(* IEC 61131-3 sources: Test-Git_ESME26/TestProgettoESME_26.fbsproj/TemplateFullProgrammingFramework_Migration.device.xml.v3^/Plc Logic.plclogic.xml.v3^/Application.application.xml.v3^/TemplateFullProgrammingFramework/Examples/ExampleDiagSources/FB_ApplicationLoggerDiagSource.fb.st^, 6 files *)

(* ---- CancelWriting.meth.st ---- *)
METHOD INTERNAL CancelWriting
VAR_INPUT
END_VAR

(* Deactivate writing if we are (for whatever reason) no longer adressed.
   May happen in case network connection with Diagnostics is disrupted or Source will be disabled *)

THIS^.diOldCmd			:= 0;
THIS^.diCmdExecState	:= 0;

(* ---- DiagQuit.meth.st ---- *)
METHOD INTERNAL DiagQuit
VAR_INPUT
END_VAR

IF THIS^.i_xEnable AND THIS^.q_xActive AND THIS^.q_etDiag <> GD.ET_Diag.Ok AND THIS^.diState = 0 THEN

	THIS^.rtrigDiagQuit(CLK := THIS^.i_xDiagQuit);
	IF THIS^.rtrigDiagQuit.Q THEN
		CancelWriting();

		THIS^.udiOwnSourceId	:= 0;

		THIS^.fbTreeWriter.FB_Init(bInitRetains := FALSE, bInCopyCode := FALSE);

		THIS^.q_xReady		:= TRUE;
		THIS^.q_etDiag		:= GD.ET_Diag.Ok;
		THIS^.q_etDiagExt	:= ET_DiagExt.WaitUntilDiagnosticsManagerReady;
		THIS^.q_sMsg		:= '';

		THIS^.diState := 10;
	END_IF

END_IF

(* ---- ExceptionDuringWriting.meth.st ---- *)
METHOD INTERNAL ExceptionDuringWriting : BOOL
VAR_INPUT
END_VAR

(* exception during writing *)
CASE THIS^.etDiagExtBufferTPL OF
	TPL.ET_DiagExt.TreeStartAlreadySuccessfullyCalled,		// FB_TreeWriter.TreeStart
	TPL.ET_DiagExt.FileIdNotSet,							// FB_TreeWriter.TreeStart
	TPL.ET_DiagExt.FileIdInvalid,							// FB_TreeWriter.TreeStart & FB_TreeWriter.NodeStart & FB_TreeWriter.Parameter & FB_TreeWriter.NodeEnd & FB_TreeWriter.TreeEnd
	TPL.ET_DiagExt.FileNotOpen,								// FB_TreeWriter.TreeStart & FB_TreeWriter.NodeStart & FB_TreeWriter.Parameter & FB_TreeWriter.NodeEnd & FB_TreeWriter.TreeEnd
	TPL.ET_DiagExt.UnexpectedFeedback,						// FB_TreeWriter.TreeStart & FB_TreeWriter.NodeStart & FB_TreeWriter.Parameter & FB_TreeWriter.NodeEnd & FB_TreeWriter.TreeEnd
	TPL.ET_DiagExt.TreeStartNotCalled,						// FB_TreeWriter.NodeStart
	TPL.ET_DiagExt.TreeStartNotSuccessfullyCalled,			// FB_TreeWriter.NodeStart
	TPL.ET_DiagExt.NoMoreNodeOpen,							// FB_TreeWriter.Parameter & FB_TreeWriter.NodeEnd
	TPL.ET_DiagExt.CallTreeStartFirst,						// FB_TreeWriter.TreeEnd
	TPL.ET_DiagExt.NodesStillOpen:							// FB_TreeWriter.TreeEnd

		SetDiagOutputs(	i_etDiag	:= GD.ET_Diag.UnexpectedProgramBehavior,
						i_etDiagExt	:= ET_DiagExt.UnexpectedFeedback,
						i_sMsg		:= SE_CTBX.FC_MultiConcat(	i_sString1	:= 'FB_TreeWriter: ',
															i_sString2	:= GD.FC_EtDiagToString(THIS^.etDiagBuffer),
															i_sString3	:= ' - ',
															i_sString4	:= TPL.FC_EtDiagExtToString(THIS^.etDiagExtBufferTPL)));
	ELSE
		SetDiagOutputs(	i_etDiag	:= GD.ET_Diag.UnexpectedProgramBehavior,
						i_etDiagExt	:= ET_DiagExt.UnexpectedFeedback,
						i_sMsg		:= SE_CTBX.FC_MultiConcat(	i_sString1	:= 'FB_TreeWriter: ',
															i_sString2	:= GD.FC_EtDiagToString(THIS^.etDiagBuffer),
															i_sString3	:= ' - ',
															i_sString4	:= TPL.FC_EtDiagExtToString(THIS^.etDiagExtBufferTPL)));

END_CASE

CancelWriting();

(* ---- SetDiagOutputs.meth.st ---- *)
METHOD INTERNAL SetDiagOutputs : BOOL
VAR_INPUT
	i_etDiag		: GD.ET_Diag;
	i_etDiagExt		: ET_DiagExt;
	i_sMsg			: STRING[80];
END_VAR

IF THIS^.q_etDiag = GD.ET_Diag.Ok OR i_etDiagExt = ET_DiagExt.Disabled THEN

	IF i_etDiag <> GD.ET_Diag.Ok OR i_etDiagExt = ET_DiagExt.Disabled THEN

		IF i_etDiag <> GD.ET_Diag.Ok THEN
			THIS^.iq_stComStructure.iq_diCmd := -THIS^.iq_stComStructure.iq_diCmd;
		END_IF

		IF i_etDiagExt = ET_DiagExt.Disabled THEN
			THIS^.q_xActive := FALSE;

			CancelWriting();
		END_IF

		THIS^.q_xReady := FALSE;
		THIS^.diState := 0;
	END_IF

	THIS^.q_etDiag		:= i_etDiag;
	THIS^.q_etDiagExt	:= i_etDiagExt;
	THIS^.q_sMsg		:= i_sMsg;
END_IF

(* ---- WriteDiagDataControl.meth.st ---- *)
METHOD INTERNAL WriteDiagDataControl : BOOL
VAR_INPUT
END_VAR

IF (THIS^.diOldCmd <> THIS^.iq_stComStructure.iq_diCmd AND THIS^.iq_stComStructure.iq_diCmd > 0) THEN
	THIS^.diOldCmd := THIS^.iq_stComStructure.iq_diCmd;

	(* new command, start execution *)
	IF THIS^.iq_stComStructure.iq_diCmd = 1 THEN
		IF (THIS^.iq_stComStructure.i_diFileId > 0) THEN
			SetDiagOutputs(	i_etDiag		:= GD.ET_Diag.Ok,
							i_etDiagExt		:= ET_DiagExt.WritingToFile,
							i_sMsg			:= '');
			THIS^.iq_stComStructure.q_lrProgress := 0.0;
			THIS^.fbTreeWriter.diFileId := THIS^.iq_stComStructure.i_diFileId;
			THIS^.diCmdExecState := 1; (* start writing to file *)
		ELSE
			(* invalid file id *)
			SetDiagOutputs(	i_etDiag		:= GD.ET_Diag.InputParameterInvalid,
							i_etDiagExt		:= ET_DiagExt.FileIdInvalid,
							i_sMsg			:= CONCAT('Invalid file Id iq_stComStructure.i_diFileId: ', TO_STRING(THIS^.iq_stComStructure.i_diFileId)));
		END_IF
	ELSE
		(* unkown cmd *)
		SetDiagOutputs(	i_etDiag		:= GD.ET_Diag.InputParameterInvalid,
						i_etDiagExt		:= ET_DiagExt.CmdUnknown,
						i_sMsg			:= CONCAT('Unknown command iq_stComStructure.diCmd: ', DINT_TO_STRING(THIS^.iq_stComStructure.iq_diCmd)));

		CancelWriting();
	END_IF
END_IF

(* ---- WriteDiagDataToFile.meth.st ---- *)
METHOD WriteDiagDataToFile
VAR_INPUT
END_VAR

TPL.FC_CanContinueWriting(iq_stCanContinueWriting := THIS^.iq_stComStructure.iq_stCanContinueWriting); (* loop as long as we can continue to write *)

WHILE (THIS^.iq_stComStructure.iq_stCanContinueWriting.xCanContinue) DO

	CASE THIS^.diCmdExecState OF
		1:	(* start writing *)
			THIS^.fbTreeWriter.TreeStart(	i_sName					:= THIS^.c_sName,
											i_sTypeName				:= THIS^.c_sTypeName,
											i_sTitleEnglish			:= 'ApplicationLogger',
											i_sTitleGerman			:= 'ApplicationLogger',
											i_uiPrintRank			:= 14,
											i_sEmptyListTextEnglish	:= 'No data available to show',
											i_sEmptyListTextGerman	:= 'Keine Daten zum Anzeigen vorhanden',
											q_etDiag				=> THIS^.etDiagBuffer,
											q_etDiagExt				=> THIS^.etDiagExtBufferTPL,
											q_sMsg					=> THIS^.sMsgBuffer);
			IF THIS^.etDiagBuffer <> GD.ET_Diag.Ok THEN
				ExceptionDuringWriting();
				EXIT;
			END_IF
			THIS^.diCmdExecState := 50;

		50:	(* Start LogEntryList *)
			THIS^.fbTreeWriter.NodeStart(	i_sName		:= 'LogEntry list',
											q_etDiag	=> etDiagBuffer,
											q_etDiagExt	=> etDiagExtBufferTPL,
											q_sMsg		=> sMsgBuffer);
			IF THIS^.etDiagBuffer <> GD.ET_Diag.Ok THEN
				ExceptionDuringWriting();
				EXIT;
			END_IF
			THIS^.udiLogEntryCount := 1;
			THIS^.udiLogEntryCountMax := 50;
			THIS^.udiLogEntryId := THIS^.fbAppLogHandler.udiFirstLogEntryId;
			THIS^.diCmdExecState := 51;

		51: (* write LogEntrys *)
			WHILE (THIS^.udiLogEntryCount < THIS^.udiLogEntryCountMax) AND (THIS^.udiLogEntryCount <= THIS^.fbAppLogHandler.udiNumberOfLogEntries) DO
				THIS^.fbTreeWriter.NodeStart(	i_sName		:= UDINT_TO_STRING(THIS^.udiLogEntryId),
												q_etDiag	=> etDiagBuffer,
												q_etDiagExt	=> etDiagExtBufferTPL,
												q_sMsg		=> sMsgBuffer);
				IF THIS^.etDiagBuffer <> GD.ET_Diag.Ok THEN
					ExceptionDuringWriting();
					RETURN;
				END_IF

					THIS^.fbAppLogHandler.GetLogEntry(	i_udiId			:= THIS^.udiLogEntryId,
														q_stLogEntry	=> THIS^.stLogEntry,
														q_etDiag		=> THIS^.etDiagBuffer,
														q_etDiagExt		=> THIS^.etDiagExtBufferAPL);
					IF (THIS^.etDiagBuffer <> GD.ET_Diag.Ok) THEN
						ExceptionDuringWriting();
						RETURN;
					END_IF

					THIS^.fbTreeWriter.Parameter(	i_sName		:= 'udiId',
													i_sValue	:= UDINT_TO_STRING(THIS^.stLogEntry.udiId),
													q_etDiag	=> etDiagBuffer,
													q_etDiagExt	=> etDiagExtBufferTPL,
													q_sMsg		=> sMsgBuffer);
					IF etDiagBuffer <> GD.ET_Diag.Ok THEN
						ExceptionDuringWriting();
						RETURN;
					END_IF

					THIS^.fbTreeWriter.Parameter(	i_sName		:= 'udiLoggerPointId',
													i_sValue	:= UDINT_TO_STRING(THIS^.stLogEntry.udiLoggerPointId),
													q_etDiag	=> etDiagBuffer,
													q_etDiagExt	=> etDiagExtBufferTPL,
													q_sMsg		=> sMsgBuffer);
					IF etDiagBuffer <> GD.ET_Diag.Ok THEN
						ExceptionDuringWriting();
						RETURN;
					END_IF
					THIS^.fbTreeWriter.Parameter(	i_sName		:= 'sMessage',
													i_sValue	:= THIS^.stLogEntry.sMessage,
													q_etDiag	=> etDiagBuffer,
													q_etDiagExt	=> etDiagExtBufferTPL,
													q_sMsg		=> sMsgBuffer);
					IF etDiagBuffer <> GD.ET_Diag.Ok THEN
						ExceptionDuringWriting();
						RETURN;
					END_IF
					THIS^.fbTreeWriter.Parameter(	i_sName		:= 'etDiag',
													i_sValue	:= GD.FC_EtDiagToString(i_etDiag := THIS^.stLogEntry.etDiag),
													q_etDiag	=> etDiagBuffer,
													q_etDiagExt	=> etDiagExtBufferTPL,
													q_sMsg		=> sMsgBuffer);
					IF etDiagBuffer <> GD.ET_Diag.Ok THEN
						ExceptionDuringWriting();
						RETURN;
					END_IF
					THIS^.fbTreeWriter.Parameter(	i_sName		:= 'udiDiagExt',
													i_sValue	:= UDINT_TO_STRING(THIS^.stLogEntry.udiDiagExt),
													q_etDiag	=> etDiagBuffer,
													q_etDiagExt	=> etDiagExtBufferTPL,
													q_sMsg		=> sMsgBuffer);
					IF etDiagBuffer <> GD.ET_Diag.Ok THEN
						ExceptionDuringWriting();
						RETURN;
					END_IF
					THIS^.fbTreeWriter.Parameter(	i_sName		:= 'dtDate',
													i_sValue	:= DATE_TO_STRING(THIS^.stLogEntry.dtDate),
													q_etDiag	=> etDiagBuffer,
													q_etDiagExt	=> etDiagExtBufferTPL,
													q_sMsg		=> sMsgBuffer);
					IF etDiagBuffer <> GD.ET_Diag.Ok THEN
						ExceptionDuringWriting();
						RETURN;
					END_IF
					THIS^.fbTreeWriter.Parameter(	i_sName		:= 'todTime',
													i_sValue	:= TOD_TO_STRING(THIS^.stLogEntry.todTime),
													q_etDiag	=> etDiagBuffer,
													q_etDiagExt	=> etDiagExtBufferTPL,
													q_sMsg		=> sMsgBuffer);
					IF etDiagBuffer <> GD.ET_Diag.Ok THEN
						ExceptionDuringWriting();
						RETURN;
					END_IF
					THIS^.fbTreeWriter.Parameter(	i_sName		:= 'etLogLevel',
													i_sValue	:= APL.FC_EtLogLevelToString(i_etLogLevel := THIS^.stLogEntry.etLogLevel),
													q_etDiag	=> etDiagBuffer,
													q_etDiagExt	=> etDiagExtBufferTPL,
													q_sMsg		=> sMsgBuffer);
					IF etDiagBuffer <> GD.ET_Diag.Ok THEN
						ExceptionDuringWriting();
						RETURN;
					END_IF

				THIS^.fbTreeWriter.NodeEnd(	q_etDiag	=> etDiagBuffer,
											q_etDiagExt	=> etDiagExtBufferTPL,
											q_sMsg		=> sMsgBuffer);
				IF THIS^.etDiagBuffer <> GD.ET_Diag.Ok THEN
					ExceptionDuringWriting();
					RETURN;
				END_IF

				THIS^.udiLogEntryCount := THIS^.udiLogEntryCount +1;
				THIS^.udiLogEntryId := THIS^.udiLogEntryId +1;
			END_WHILE
			THIS^.udiLogEntryCountMax := THIS^.udiLogEntryCountMax + 50;
			IF (THIS^.udiLogEntryCount > THIS^.fbAppLogHandler.udiNumberOfLogEntries) THEN
				THIS^.fbTreeWriter.NodeEnd(	q_etDiag	=> etDiagBuffer,
											q_etDiagExt	=> etDiagExtBufferTPL,
											q_sMsg		=> sMsgBuffer);
				IF THIS^.etDiagBuffer <> GD.ET_Diag.Ok THEN
					ExceptionDuringWriting();
					EXIT;
				END_IF
				THIS^.diCmdExecState := 60;
			END_IF

		60: (* Start LoggerPoint list *)
			THIS^.fbTreeWriter.NodeStart(	i_sName		:= 'LoggerPoint list',
											q_etDiag	=> etDiagBuffer,
											q_etDiagExt	=> etDiagExtBufferTPL,
											q_sMsg		=> sMsgBuffer);
			IF THIS^.etDiagBuffer <> GD.ET_Diag.Ok THEN
				ExceptionDuringWriting();
				EXIT;
			END_IF
			THIS^.udiLoggerPointCount := 1;
			THIS^.udiLoggerPointCountMax := 50;
			THIS^.diCmdExecState := 61;

		61: (* write LoggerPoint list *)
			WHILE (THIS^.udiLoggerPointCount < THIS^.udiLoggerPointCountMax) AND (THIS^.udiLoggerPointCount <= THIS^.fbAppLogHandler.udiNumberOfLoggerPoints) DO
				THIS^.fbTreeWriter.NodeStart(	i_sName		:= UDINT_TO_STRING(THIS^.udiLoggerPointCount),
												q_etDiag	=> etDiagBuffer,
												q_etDiagExt	=> etDiagExtBufferTPL,
												q_sMsg		=> sMsgBuffer);
				IF THIS^.etDiagBuffer <> GD.ET_Diag.Ok THEN
					ExceptionDuringWriting();
					RETURN;
				END_IF

					THIS^.fbAppLogHandler.GetLoggerPoint(	i_udiId			:= THIS^.udiLoggerPointCount,
															q_ifLoggerPoint	=> THIS^.ifLoggerPoint,
															q_etDiag		=> THIS^.etDiagBuffer,
															q_etDiagExt		=> THIS^.etDiagExtBufferAPL);
					IF (THIS^.etDiagBuffer <> GD.ET_Diag.Ok) THEN
						ExceptionDuringWriting();
						RETURN;
					END_IF

					THIS^.fbTreeWriter.Parameter(	i_sName		:= 'udiId',
													i_sValue	:= UDINT_TO_STRING(THIS^.ifLoggerPoint.udiId),
													q_etDiag	=> etDiagBuffer,
													q_etDiagExt	=> etDiagExtBufferTPL,
													q_sMsg		=> sMsgBuffer);
					IF etDiagBuffer <> GD.ET_Diag.Ok THEN
						ExceptionDuringWriting();
						RETURN;
					END_IF
					THIS^.fbTreeWriter.Parameter(	i_sName		:= 'udiParentId',
													i_sValue	:= UDINT_TO_STRING(THIS^.ifLoggerPoint.udiParentId),
													q_etDiag	=> etDiagBuffer,
													q_etDiagExt	=> etDiagExtBufferTPL,
													q_sMsg		=> sMsgBuffer);
					IF etDiagBuffer <> GD.ET_Diag.Ok THEN
						ExceptionDuringWriting();
						RETURN;
					END_IF
					THIS^.fbTreeWriter.Parameter(	i_sName		:= 'sName',
													i_sValue	:= THIS^.ifLoggerPoint.sName,
													q_etDiag	=> etDiagBuffer,
													q_etDiagExt	=> etDiagExtBufferTPL,
													q_sMsg		=> sMsgBuffer);
					IF etDiagBuffer <> GD.ET_Diag.Ok THEN
						ExceptionDuringWriting();
						RETURN;
					END_IF
					THIS^.fbTreeWriter.Parameter(	i_sName		:= 'sType',
													i_sValue	:= THIS^.ifLoggerPoint.sType,
													q_etDiag	=> etDiagBuffer,
													q_etDiagExt	=> etDiagExtBufferTPL,
													q_sMsg		=> sMsgBuffer);
					IF etDiagBuffer <> GD.ET_Diag.Ok THEN
						ExceptionDuringWriting();
						RETURN;
					END_IF
					THIS^.fbTreeWriter.Parameter(	i_sName		:= 'sSource',
													i_sValue	:= THIS^.ifLoggerPoint.sSource,
													q_etDiag	=> etDiagBuffer,
													q_etDiagExt	=> etDiagExtBufferTPL,
													q_sMsg		=> sMsgBuffer);
					IF etDiagBuffer <> GD.ET_Diag.Ok THEN
						ExceptionDuringWriting();
						RETURN;
					END_IF
					THIS^.fbTreeWriter.Parameter(	i_sName		:= 'etLogLevel',
													i_sValue	:= APL.FC_EtLogLevelToString(i_etLogLevel := THIS^.ifLoggerPoint.etLogLevel),
													q_etDiag	=> etDiagBuffer,
													q_etDiagExt	=> etDiagExtBufferTPL,
													q_sMsg		=> sMsgBuffer);
					IF etDiagBuffer <> GD.ET_Diag.Ok THEN
						ExceptionDuringWriting();
						RETURN;
					END_IF

				THIS^.fbTreeWriter.NodeEnd(	q_etDiag	=> etDiagBuffer,
											q_etDiagExt	=> etDiagExtBufferTPL,
											q_sMsg		=> sMsgBuffer);
				IF THIS^.etDiagBuffer <> GD.ET_Diag.Ok THEN
					ExceptionDuringWriting();
					RETURN;
				END_IF

				THIS^.udiLoggerPointCount := THIS^.udiLoggerPointCount +1;
			END_WHILE
			THIS^.udiLoggerPointCountMax := THIS^.udiLoggerPointCountMax + 50;
			IF (THIS^.udiLoggerPointCount > THIS^.fbAppLogHandler.udiNumberOfLoggerPoints) THEN
				THIS^.fbTreeWriter.NodeEnd(	q_etDiag	=> etDiagBuffer,
											q_etDiagExt	=> etDiagExtBufferTPL,
											q_sMsg		=> sMsgBuffer);
				IF THIS^.etDiagBuffer <> GD.ET_Diag.Ok THEN
					ExceptionDuringWriting();
					EXIT;
				END_IF
				THIS^.diCmdExecState := 70;
			END_IF

		70:
			(* library versions *)
			THIS^.fbTreeWriter.NodeStart(	i_sName		:= 'LibraryVersions',
											q_etDiag	=> THIS^.etDiagBuffer,
											q_etDiagExt	=> THIS^.etDiagExtBufferTPL,
											q_sMsg		=> THIS^.sMsgBuffer);
			IF THIS^.etDiagBuffer <> GD.ET_Diag.Ok THEN
				ExceptionDuringWriting();
				EXIT;
			END_IF

				THIS^.fbTreeWriter.Parameter(	i_sName		:= 'ApplicationLogger',
												i_sValue	:= APL.Gc_sLibraryVersion,
												q_etDiag	=> THIS^.etDiagBuffer,
												q_etDiagExt	=> THIS^.etDiagExtBufferTPL,
												q_sMsg		=> THIS^.sMsgBuffer);
				IF THIS^.etDiagBuffer <> GD.ET_Diag.Ok THEN
					ExceptionDuringWriting();
					EXIT;
				END_IF

				THIS^.fbTreeWriter.Parameter(	i_sName		:= 'GlobalDiagnostics',
												i_sValue	:= GD.Gc_sLibraryVersion,
												q_etDiag	=> THIS^.etDiagBuffer,
												q_etDiagExt	=> THIS^.etDiagExtBufferTPL,
												q_sMsg		=> THIS^.sMsgBuffer);
				IF THIS^.etDiagBuffer <> GD.ET_Diag.Ok THEN
					ExceptionDuringWriting();
					EXIT;
				END_IF

			THIS^.fbTreeWriter.NodeEnd(	q_etDiag	=> THIS^.etDiagBuffer,
										q_etDiagExt	=> THIS^.etDiagExtBufferTPL,
										q_sMsg		=> THIS^.sMsgBuffer);
			IF THIS^.etDiagBuffer <> GD.ET_Diag.Ok THEN
				ExceptionDuringWriting();
				EXIT;
			END_IF

			THIS^.fbTreeWriter.TreeEnd(	q_etDiag	=> THIS^.etDiagBuffer,
										q_etDiagExt	=> THIS^.etDiagExtBufferTPL,
										q_sMsg		=> THIS^.sMsgBuffer);
			IF THIS^.etDiagBuffer <> GD.ET_Diag.Ok THEN
				ExceptionDuringWriting();
				EXIT;
			END_IF
			(* done *)

			(* signal command execution *)
			THIS^.iq_stComStructure.iq_diCmd := 0;

			SetDiagOutputs(	i_etDiag	:= GD.ET_Diag.Ok,
							i_etDiagExt	:= ET_DiagExt.DataSuccessfullyWritten,
							i_sMsg		:= '');

			THIS^.diCmdExecState := 0;
			EXIT; (* exit the while loop *)
		ELSE
			ExceptionDuringWriting();
			EXIT;
	END_CASE
END_WHILE
